Staubli VAL3: HMI_FrameSet.pjx

--- HMI_FrameSet.pjx ---
Parameters version=s8.15.3Cs9_BS3337 stackSize=5000 millimeterUnit=true
Program file=bind.pgx
Program file=computeFrame.pgx
Program file=getIndex.pgx
Program file=main.pgx
Program file=modifyFrame.pgx
Program file=movePoint.pgx
Program file=nmbValue.pgx
Program file=onStart.pgx
Program file=refreshList.pgx
Program file=renameFrame.pgx
Program file=renameTool.pgx
Program file=setTool.pgx
Program file=start.pgx
Program file=stop.pgx
Program file=teachPoint.pgx
Program file=wizard.pgx
Data file=HMI_FrameSet.dtx
Library alias=util path=Disk://HMI_cs9/HMI_util/HMI_util.pjx
Library alias=savedata path=Disk://source/saveData/saveData.pjx

--- HMI_FrameSet.dtx ---
mdesc mNomSpeed = {accel=25, vel=50, decel=25, leave=0, reach=0, blend=off}
string sFrameList
string sToolList
string sSelFrame
string sSelTool
bool bBool[6]
bool bBack
public num nTool[6]
bool bModifyTool
bool bCancelTool
num nFrame[6]
bool bModifyFrame
bool bCancelFrame
string sUsingTool
string sUsingFrame
num nNmbValue[6]
num nWizardStep
bool bPrevious
bool bTeach
bool bMove
bool bNext
string sLastTool
tool tUsingTool = {fatherId=flange[0]}
string sTitle
num _nTool

--- main.pgx ---
public program main()
  local bool l_bRefresh
  local num l_nPoint
  local bool l_bExit
begin
  do
    if util:sPage!="frame"
      util:sPage="frame"
      call onStart()
      call bind()
      call util:loadingPage()
      userPage(util:sPage)
      delay(0.5)
    endIf
    //button
    if bBool[1]
      bBool[1]=false
      call getIndex(sSelFrame,l_nPoint)
      if l_nPoint!=0
        call wizard(l_nPoint)
      else
        userPageAlert("0号frame不可修改")
      endIf
    elseIf bBool[2]
      bBool[2]=false
      //modify frame
      call getIndex(sSelFrame,l_nPoint)
      if l_nPoint!=0
        call modifyFrame(l_nPoint)
      else
        userPageAlert("0号frame不可修改")
      endIf
    elseIf bBool[3]
      bBool[3]=false
      //重命名frame
      call getIndex(sSelFrame,l_nPoint)
      if l_nPoint!=0
        call renameFrame(l_nPoint)
      else
        userPageAlert("0号frame不可修改")
      endIf
      l_bRefresh=true
    elseIf bBool[4]
      bBool[4]=false
      //modify tool
      call getIndex(sSelTool,l_nPoint)
      if l_nPoint!=0
        call setTool(l_nPoint)
      else
        userPageAlert("0号tool不可修改")
      endIf
    elseIf bBool[5]
      bBool[5]=false
      //重命名tool
      call getIndex(sSelTool,l_nPoint)
      if l_nPoint!=0
        call renameTool(l_nPoint)
      else
        userPageAlert("0号tool不可修改")
      endIf
      l_bRefresh=true
    elseIf bBack
      bBack=false
      l_bExit=true

    endIf

    //refresh
    if l_bRefresh
      l_bRefresh=false
      call refreshList()
    endIf



    delay(0)
  until l_bExit==true
end

--- start.pgx ---
program start()
begin
end

--- bind.pgx ---
program bind()
  local string l_sbtn
  local num l_i
begin
  userPageBind("frame","lst1","options",sFrameList,size(sFrameList),"r")
  userPageBind("frame","lst2","options",sToolList,size(sToolList),"r")
  userPageBind("frame","lst1","value",sSelFrame,1,"rw")
  userPageBind("frame","lst2","value",sSelTool,1,"rw")
  //button
  for l_i =1 to 5
    l_sbtn="btn"+toString("",l_i)
    userPageBindClick("frame",l_sbtn,bBool[l_i],true)
  endFor
  userPageBindClick("frame","btnback",bBack,true)
end

--- computeFrame.pgx ---
program computeFrame(num x_nIndex)
  local num l_nResult
begin

  l_nResult= setFrame(savedata:fFrameItem[x_nIndex].pPointRx[0],savedata:fFrameItem[x_nIndex].pPointRx[1],savedata:fFrameItem[x_nIndex].pPointRx[2],savedata:fFrameItem[x_nIndex].fFrame)
  popUpMsg("坐标系计算完成")
  savedata:libSave()
  delay(0.1)
  if l_nResult<0
    userPageAlert("坐标系示教不成功！请重新示教")
  endIf

end

--- getIndex.pgx ---
public program getIndex(string x_sKey, num& x_nIndex)
  local bool l_bResult
  local num l_nIndex
begin
  toNum(x_sKey,l_nIndex,l_bResult)
  if l_bResult
    x_nIndex=l_nIndex
  else
    x_nIndex=-1
    userPageAlert("未选择有效项目！")
  endIf
end

--- modifyFrame.pgx ---
program modifyFrame(num x_nIndex)
  local bool l_bExit
  local num l_i
  local string l_sNmb
begin
  do
    if util:sPage!="frameSetting"
      util:sPage="frameSetting"

      nFrame[0]=savedata:fFrameItem[x_nIndex].fFrame.trsf.x
      nFrame[1]=savedata:fFrameItem[x_nIndex].fFrame.trsf.y
      nFrame[2]=savedata:fFrameItem[x_nIndex].fFrame.trsf.z
      nFrame[3]=savedata:fFrameItem[x_nIndex].fFrame.trsf.rx
      nFrame[4]=savedata:fFrameItem[x_nIndex].fFrame.trsf.ry
      nFrame[5]=savedata:fFrameItem[x_nIndex].fFrame.trsf.rz
      for l_i = 0 to 5
        l_sNmb="nmb"+toString("",l_i+1)
        userPageBind("frameSetting",l_sNmb,"value",nFrame[l_i],1,"rw")
      endFor
      userPageBindClick("frameSetting","btn1",bModifyFrame,true)
      userPageBindClick("frameSetting","btn2",bCancelFrame,true)
      userPage(util:sPage)
      delay(0.5)
    endIf

    if bModifyFrame
      bModifyFrame=false
      savedata:fFrameItem[x_nIndex].fFrame.trsf.x=nFrame[0]
      savedata:fFrameItem[x_nIndex].fFrame.trsf.y=nFrame[1]
      savedata:fFrameItem[x_nIndex].fFrame.trsf.z=nFrame[2]
      savedata:fFrameItem[x_nIndex].fFrame.trsf.rx=nFrame[3]
      savedata:fFrameItem[x_nIndex].fFrame.trsf.ry=nFrame[4]
      savedata:fFrameItem[x_nIndex].fFrame.trsf.rz=nFrame[5]
      savedata:libSave()
      delay(0.1)
       l_bExit=true
    elseIf bCancelFrame
      bCancelFrame=false
      l_bExit=true
    endIf
    delay(0)
  until l_bExit==true
end

--- movePoint.pgx ---
program movePoint(num x_nStep, num x_nIndex)
  local bool l_bResult
begin
  //   l_bResult=userPageConfirm("是否移动到该点位？")
  //  if l_bResult
  resetMotion()
  $jogMode(0)
  switch x_nStep
    case 0
      movel(savedata:fFrameItem[x_nIndex].pPointRx[0],tUsingTool,mNomSpeed)
    break
    case 1
      movel(savedata:fFrameItem[x_nIndex].pPointRx[1],tUsingTool,mNomSpeed)
    break
    case 2
      movel(savedata:fFrameItem[x_nIndex].pPointRx[2],tUsingTool,mNomSpeed)
    break
  endSwitch
  //  endIf
end

--- nmbValue.pgx ---
program nmbValue(num x_nStep, num x_nIndex)
  local trsf l_trsf
  local num l_nResult
begin
  switch x_nStep

    case 0
      l_trsf=savedata:fFrameItem[x_nIndex].pPointRx[0].trsf
      sUsingFrame=savedata:fFrameItem[x_nIndex].sName+" 坐标系O点"
      nNmbValue[0]=l_trsf.x
      nNmbValue[1]=l_trsf.y
      nNmbValue[2]=l_trsf.z
      nNmbValue[3]=l_trsf.rx
      nNmbValue[4]=l_trsf.ry
      nNmbValue[5]=l_trsf.rz
    break
    case 1
      l_trsf=savedata:fFrameItem[x_nIndex].pPointRx[1].trsf
      sUsingFrame=savedata:fFrameItem[x_nIndex].sName+" 坐标系X点"
      nNmbValue[0]=l_trsf.x
      nNmbValue[1]=l_trsf.y
      nNmbValue[2]=l_trsf.z
      nNmbValue[3]=l_trsf.rx
      nNmbValue[4]=l_trsf.ry
      nNmbValue[5]=l_trsf.rz
    break
    case 2
      l_trsf=savedata:fFrameItem[x_nIndex].pPointRx[2].trsf
      sUsingFrame=savedata:fFrameItem[x_nIndex].sName+" 坐标系Y点"
      nNmbValue[0]=l_trsf.x
      nNmbValue[1]=l_trsf.y
      nNmbValue[2]=l_trsf.z
      nNmbValue[3]=l_trsf.rx
      nNmbValue[4]=l_trsf.ry
      nNmbValue[5]=l_trsf.rz
    break


  endSwitch




end

--- onStart.pgx ---
program onStart()
  local num l_nSize
  local num l_i
begin
  l_nSize=size(savedata:fFrameItem)
  resize(sFrameList,1,l_nSize)
  l_nSize=size(savedata:tToolItem)
  resize(sToolList,1,l_nSize)

  for l_i = 0 to size(sFrameList)-1
    sFrameList[l_i]=toString("",l_i)+","+savedata:fFrameItem[l_i].sName
  endFor

  for l_i = 0 to size(sToolList)-1
    sToolList[l_i]=toString("",l_i)+","+savedata:tToolItem[l_i].sName
  endFor

  sSelFrame=sFrameList[0]
  sSelTool=sToolList[0]

end

--- refreshList.pgx ---
program refreshList()
  local num l_i
begin
  for l_i = 0 to size(sFrameList)-1
    sFrameList[l_i]=toString("",l_i)+","+savedata:fFrameItem[l_i].sName
  endFor

  for l_i = 0 to size(sToolList)-1
    sToolList[l_i]=toString("",l_i)+","+savedata:tToolItem[l_i].sName
  endFor
end

--- renameFrame.pgx ---
program renameFrame(num x_nIndex)
  local string l_sName
  local bool l_bResult
begin
  l_bResult=userPagePrompt("请输入新的名称：",l_sName)
  if l_bResult
    savedata:fFrameItem[x_nIndex].sName=l_sName
    savedata:libSave()
    delay(0.1)
  endIf
end

--- renameTool.pgx ---
program renameTool(num x_nIndex)
  local string l_sName
  local bool l_bResult
begin
  l_bResult=userPagePrompt("请输入新的名称：",l_sName)
  if l_bResult
    savedata:tToolItem[x_nIndex].sName=l_sName
    savedata:libSave()
    delay(0.1)
  endIf
end

--- setTool.pgx ---
program setTool(num x_nIndex)
  local bool l_bExit
  local num l_nUsingTool
  local string l_sNmb
  local num l_i
begin
  do
    if util:sPage!="toolSetting"
      util:sPage="toolSetting"
      l_nUsingTool=x_nIndex
      nTool[0]=savedata:tToolItem[x_nIndex].tTool.trsf.x
      nTool[1]=savedata:tToolItem[x_nIndex].tTool.trsf.y
      nTool[2]=savedata:tToolItem[x_nIndex].tTool.trsf.z
      nTool[3]=savedata:tToolItem[x_nIndex].tTool.trsf.rx
      nTool[4]=savedata:tToolItem[x_nIndex].tTool.trsf.ry
      nTool[5]=savedata:tToolItem[x_nIndex].tTool.trsf.rz
      for l_i = 0 to 5
        l_sNmb="nmb"+toString("",l_i+1)
        userPageBind("toolSetting",l_sNmb,"value",nTool[l_i],1,"rw")
      endFor
      userPageBindClick("toolSetting","btn1",bModifyTool,true)
      userPageBindClick("toolSetting","btn2",bCancelTool,true)
      userPageBind("toolSetting","lbltitle","innerHTML",sTitle,1,"r")
      sTitle="设定工具："+toString("",l_nUsingTool)
      userPage(util:sPage)
      delay(0.5)
      //l_bExit=true
    endIf

    if bModifyTool
      bModifyTool=false
      savedata:tToolItem[x_nIndex].tTool.trsf.x=nTool[0]
      savedata:tToolItem[x_nIndex].tTool.trsf.y=nTool[1]
      savedata:tToolItem[x_nIndex].tTool.trsf.z=nTool[2]
      savedata:tToolItem[x_nIndex].tTool.trsf.rx=nTool[3]
      savedata:tToolItem[x_nIndex].tTool.trsf.ry=nTool[4]
      savedata:tToolItem[x_nIndex].tTool.trsf.rz=nTool[5]
      savedata:libSave()
      l_bExit=true
      delay(0.1)
    elseIf bCancelTool
      bCancelTool=false
      l_bExit=true
    endIf
    delay(0)
  until l_bExit==true
end

--- stop.pgx ---
program stop()
begin
end

--- teachPoint.pgx ---
program teachPoint(num x_nStep, num x_nIndex)
  local bool l_bResult
begin
  l_bResult=userPageConfirm("是否记录该点位？")
  if l_bResult
    switch x_nStep
      case 0
        savedata:fFrameItem[x_nIndex].pPointRx[0]=here(tUsingTool,world)
      break
      case 1
        savedata:fFrameItem[x_nIndex].pPointRx[1]=here(tUsingTool,world)
      break
      case 2
        savedata:fFrameItem[x_nIndex].pPointRx[2]=here(tUsingTool,world)
      break

    endSwitch
  endIf
end

--- wizard.pgx ---
program wizard(num x_nIndex)
  local bool l_bExit
  local string l_snmb
  local bool l_bResult
  local num l_nTool
  local tool l_tTool
  local bool l_bRefresh
  local num l_i
begin
  do
    if util:sPage!="Wizard"
      util:sPage="Wizard"
      sUsingTool=""
      sLastTool=""
      nWizardStep=0
      sUsingFrame=savedata:fFrameItem[x_nIndex].sName+" 坐标系O点"
      call nmbValue(nWizardStep,x_nIndex)
      userPageBind("Wizard","cbx1","options",sToolList,size(sToolList),"r")
      userPageBind("Wizard","cbx1","value",sUsingTool,1,"rw")
      userPageBind("Wizard","lbl2","innerHTML",sUsingFrame,1,"r")
      for l_i = 0 to size(nNmbValue)-1
        l_snmb="nmb"+toString("",l_i+1)
        userPageBind("Wizard",l_snmb,"value",nNmbValue[l_i],1,"rw")
      endFor
      userPageBindClick("Wizard","btn4",bPrevious,true)
      userPageBindClick("Wizard","btn1",bTeach,true)
      userPageBindClick("Wizard","btn3",bMove,true)
      userPageBindClick("Wizard","btn2",bNext,true)
      userPage(util:sPage)
      delay(0.5)
      _nTool=0
    endIf

    if sUsingTool!=sLastTool
      sLastTool=sUsingTool
      toNum(sLastTool,_nTool,l_bResult)
      call savedata:getTool(_nTool,tUsingTool)
      $jogContext(tUsingTool,world,0)
    endIf

    if bPrevious
      bPrevious=false
      nWizardStep=nWizardStep-1
      if nWizardStep<0
        l_bExit=true
      endIf
      l_bRefresh=true
    elseIf bTeach
      bTeach=false
      if sUsingTool!=""
        call teachPoint(nWizardStep,x_nIndex)
      else
        userPageAlert("选择有效的tool！")
      endIf
      l_bRefresh=true
    elseIf bMove
      bMove=false
      if sUsingTool!=""
        call movePoint(nWizardStep,x_nIndex)
      else
        userPageAlert("选择有效的tool！")
      endIf


    elseIf bNext
      bNext=false
      nWizardStep=nWizardStep+1
      if nWizardStep>2
        call computeFrame(x_nIndex)
        l_bExit=true
      endIf
      l_bRefresh=true
    endIf

    if l_bRefresh
      l_bRefresh=false
      if nWizardStep>0
        userPageSet("Wizard","cbx1","disabled",true)
      else
        userPageSet("Wizard","cbx1","disabled",false)
      endIf

      call nmbValue(nWizardStep,x_nIndex)
    endIf
    //jogmode
    call util:jogMode(_nTool,0)
    delay(0)
  until l_bExit==true
  resetMotion()
end
